(* IEC 61131-3 sources: plc-iiot-stack/src/POUs/Iiot/F_IiotIsName, 2 files *)

(* ---- F_IiotIsName.decl.st ---- *)
// Назначение: уровень топика по шаблону: первая — буква (только заглавная при xUpperOnly), дальше
//             буквы, цифры и _ (буквы только заглавные при xUpperOnly), длина 1..iMaxLen. Устройство:
//             [A-Z][A-Z0-9_]{0,15}; команда: [A-Za-z][A-Za-z0-9_]{0,31}.
// Автор:      kr0nsch
// Версия:     0.1.0
// Документ:   docs/plc_mqtt.md, раздел «Топики»
FUNCTION F_IiotIsName : BOOL
VAR_INPUT
    sText : STRING(GVL_Const.IIOT_LEVEL_LEN);
    iMaxLen : INT;
    xUpperOnly : BOOL;
END_VAR
VAR
    iLen : INT;
    iIdx : INT;
    bCh : BYTE;
    xUpper : BOOL;
    xLower : BOOL;
    xDigit : BOOL;
END_VAR

(* ---- F_IiotIsName.impl.st ---- *)
iLen := LEN(sText);
IF iLen < 1 OR iLen > iMaxLen THEN
    RETURN;
END_IF
FOR iIdx := 0 TO iLen - 1 DO
    bCh := sText[iIdx];
    xUpper := bCh >= GVL_Const.ASCII_UPPER_A AND bCh <= GVL_Const.ASCII_UPPER_Z;
    xLower := bCh >= GVL_Const.ASCII_LOWER_A AND bCh <= GVL_Const.ASCII_LOWER_Z AND NOT xUpperOnly;
    xDigit := bCh >= GVL_Const.ASCII_ZERO AND bCh <= GVL_Const.ASCII_NINE;
    IF iIdx = 0 THEN
        IF NOT (xUpper OR xLower) THEN
            RETURN;
        END_IF
    ELSIF NOT (xUpper OR xLower OR xDigit OR bCh = GVL_Const.ASCII_UNDERSCORE) THEN
        RETURN;
    END_IF
END_FOR
F_IiotIsName := TRUE;
